SUBAPPLICATION Uebung_OPC_L03_AX (* Wie Training_03, aber lokal und ohne VT: Input_I1 ruft die Toggle-Methode per CALL_METHOD an localhost auf, Output_Q2 zeigt den Zustand *)
  (* Standard: 61499-2; Description: Copyright (c) 2026 Meisterschulen am Ostbahnhof This program and the accompanying materials are made available under the terms of the Eclipse Public License 2.0 which is available at https://www.eclipse.org/legal/epl-2.0/ SPDX-License-Identifier: EPL-2.0 *)
  (* Version 1.0, 2026-10-18, Franz Höpfinger, Meisterschulen am Ostbahnhof, OPC-UA lokal auf einem Geraet (Meins/04_OPC_UA) *)
  PACKAGE Meins::OPC_UA_Lokal;
  IMPORT Meins::OPC_UA_Lokal::const::OpcUaLokal::L03_FF1_TRIGGER_CALL;
  IMPORT Meins::OPC_UA_Lokal::const::OpcUaLokal::L03_FF1_STATE_READ;
  IMPORT Meins::OPC_UA_Lokal::const::OpcUaLokal::L03_FF1_TRIGGER_METHOD;
  IMPORT Meins::OPC_UA_Lokal::const::OpcUaLokal::L03_FF1_STATE_WRITE;
  IMPORT logiBUS::io::DI::logiBUS_DI::Input_I1;
  IMPORT logiBUS::io::DQ::logiBUS_DO::Output_Q1;
  IMPORT logiBUS::io::DQ::logiBUS_DO::Output_Q2;
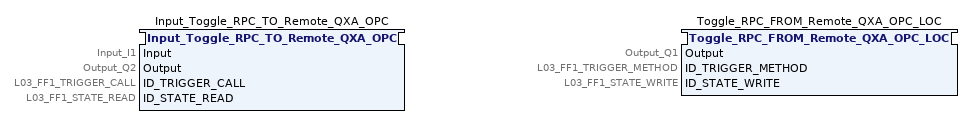
  SUBAPPS
    Input_Toggle_RPC_TO_Remote_QXA_OPC : MyLib::sys::Input_Toggle_RPC_TO_Remote_QXA_OPC(Input := Input_I1, Output := Output_Q2, ID_TRIGGER_CALL := L03_FF1_TRIGGER_CALL, ID_STATE_READ := L03_FF1_STATE_READ);
    Toggle_RPC_FROM_Remote_QXA_OPC_LOC : MyLib::sys::Toggle_RPC_FROM_Remote_QXA_OPC_LOC(Output := Output_Q1, ID_TRIGGER_METHOD := L03_FF1_TRIGGER_METHOD, ID_STATE_WRITE := L03_FF1_STATE_WRITE);
  END_SUBAPPS
END_SUBAPPLICATION
